(* IEC 61131-3 sources: trust-platform/examples/OSCAT/cold_storage_alarm/non-oop/src, 3 files *)

(* ---- Configuration.st ---- *)
CONFIGURATION ColdStorageAlarmClassicConfiguration
RESOURCE Cpu0 ON PLC
    TASK MainTask (INTERVAL := T#100ms, PRIORITY := 1);
    PROGRAM Main WITH MainTask : Main;
END_RESOURCE
END_CONFIGURATION

(* ---- Main.st ---- *)
PROGRAM Main
VAR
    TemperatureConversion : TEMPERATURE;
    DoorAlarm : HYST;
    ChamberCelsius : REAL := REAL#0.0 - REAL#16.0;
    ChamberKelvin : REAL;
    AlarmActive : BOOL;
END_VAR

TemperatureConversion(C := ChamberCelsius);
DoorAlarm(
    In := ChamberCelsius,
    HIGH_LIMIT := REAL#0.0 - REAL#18.0,
    LOW_LIMIT := REAL#0.0 - REAL#30.0
);
ChamberKelvin := TemperatureConversion.YK;
AlarmActive := DoorAlarm.Q;
END_PROGRAM

(* ---- Tests.st ---- *)
TEST_PROGRAM ColdStorageAlarmClassicDetectsWarmChamber
VAR
    TemperatureConversion : TEMPERATURE;
    DoorAlarm : HYST;
END_VAR

TemperatureConversion(C := REAL#0.0 - REAL#16.0);
DoorAlarm(
    In := REAL#0.0 - REAL#16.0,
    HIGH_LIMIT := REAL#0.0 - REAL#18.0,
    LOW_LIMIT := REAL#0.0 - REAL#30.0
);

ASSERT_NEAR(EXPECTED := REAL#257.15, ACTUAL := TemperatureConversion.YK, DELTA := REAL#0.01);
ASSERT_TRUE(IN := DoorAlarm.Q);
END_TEST_PROGRAM
